Fanuc KAREL source: KT00910.KL

PROGRAM KT00910
%NOLOCKGROUP
%ENVIRONMENT VECTR
VAR
  P1: XYZWPREXT
  P2: XYZWPREXT
  OUT: VECTOR
BEGIN
  P1.X = 1.0
  P2.Y = 2.0
  P1.X = 1.0
  P2.Y = 2.0
  OUT = ORIENT(P1)
END KT00910
